(* IEC 61131-3 sources: JingjiangMoonbox/Application/Application/任务列表/TensionTask/张力控制/收放牵/张力控制, 5 files *)

(* ---- KS_FB_CalcGirthByVel_IfOf.st ---- *)
(*@CES
Name=KS_FB_CalcGirthByVel_IfOf
Type=FunctionBlock
TypeGuid=6f9dac99-8de1-4efc-8465-68ac443b7d08
Guid=2b108746-d302-40a1-8059-c5776d7629bb
HasDeclaration=True
HasImplementation=True
*)
{DECLARATION}
FUNCTION_BLOCK KS_FB_CalcGirthByVel_IfOf
VAR_INPUT
	i_xEn: BOOL;
	i_xCalcGirthEn:BOOL;(**)
	i_rVel_Film:REAL;(*料膜速度*)
	i_iCycleTime_Plc:INT;(*程序执行周期*)
	i_rAnalogLimit:REAL;(*模拟量的限值*)
	i_rUsingGirth:REAL;(*使用的周长值*)
	i_rAnalogSumLimit:REAL;(*模拟量累计值的限值*)
	i_rAxisVel_Cur:REAL;(*当前轴速度*)
	i_rAi_Swing: REAL; (*摆臂当前值*)
END_VAR
VAR_OUTPUT
	o_xEno:BOOL;
	o_iErNo: INT;
	o_xGirthCaled:BOOL;(*周长计算完成了~*)
	o_rGirth:REAL;(*计算出来的周长值*)
END_VAR
VAR
	rAver_CurrentVel: REAL;
	rCurrentVelSum:LREAL;(*当前速度累计值*)
	rAnalogSum: REAL; (*当前模拟量累计值*)
	iCycleCount: INT;
	arDataFifo:ARRAY [1..2,1..c_iArrNum] OF REAL;(*用来存放每个周期速度以及模拟量的值。一维数组代表速度值，二维数组代表模拟量值*)
	xArrInited: BOOL;		(*数组初始化完成*)
	iDelayCount: INT;
	iN: INT;
	xAnalogValue: BOOL;(*放牵模拟量有效*)
	iLastIndex: INT;
END_VAR
VAR CONSTANT
	c_iArrNum:INT:=300;(*数组大小暂定为100个 按20ms周期算就是2s的数据*)
								(*2019.7.25.125733 将计算周期拉长了！|Liu.yt*)
END_VAR
{IMPLEMENTATION}
o_xEno:= i_xEn;
o_iErNo:= 0;
IF i_xEn THEN

	o_xGirthCaled:=FALSE;(*该标志只有效一个周期*)
	o_rGirth:=0;
	rAver_CurrentVel:=0;
	rCurrentVelSum:=0;
	rAnalogSum:=0;

	IF i_xCalcGirthEn  THEN(*使能计算周长功能*)

		(*保存一定时间的速度值，用来进行平均速度计算。时间暂定为2s*)
		iCycleCount:=iCycleCount+1;(*计数+1*)
		IF iCycleCount>c_iArrNum THEN(*循环存储*)
			iCycleCount:=1;
		END_IF
		arDataFifo[1,iCycleCount]:=i_rAxisVel_Cur;(*速度值*)
		arDataFifo[2,iCycleCount]:=i_rAi_Swing;(*模拟量值*)

		(*周长计算*)
		IF iCycleCount>=c_iArrNum OR xArrInited THEN (*累计足够次数的速度值*)

			xArrInited:=TRUE;
			iDelayCount:=iDelayCount+1;
		(*计算模拟量累计值和速度累计值*)
			FOR iN:=1 TO c_iArrNum BY 1 DO
				rCurrentVelSum:=rCurrentVelSum+arDataFifo[1,iN];
				IF ABS(arDataFifo[2,iN])>i_rAnalogLimit AND iDelayCount<=500 THEN(*累计的这段时间里的模拟量值必须都小于等于模拟量限值才有效
												iDelayCount 是用来保证在极端情况下不能满足条件也可以进入计算逻辑*)
					rAnalogSum:=i_rAnalogSumLimit+1;(*给模拟量累计值一个大于模拟量累计限值的值，这样我们在下面的判断中则会认为无效*)
					xAnalogValue:=FALSE;
					EXIT;
				ELSE
					xAnalogValue:=TRUE;
					rAnalogSum:=rAnalogSum+arDataFifo[2,iN];
				END_IF
			END_FOR

			iLastIndex:=(iCycleCount+1) MOD c_iArrNum;

			IF ABS((arDataFifo[2,iCycleCount])-(arDataFifo[2,iLastIndex])) >0.005 OR NOT  xAnalogValue THEN(*模拟量2S的变化量超过范围，则认为无效*);
			ELSE(*模拟量累计值在一定范围内求取速度平均值*)
				rAver_CurrentVel:=rCurrentVelSum/INT_TO_REAL(c_iArrNum);
			END_IF
		END_IF

		IF rAver_CurrentVel<>0 AND i_rVel_Film<>0 THEN (*平均速度不等于0 我们认为已经计算出了满足条件的平均速度值*)
			o_rGirth:=i_rVel_Film*i_rUsingGirth/rAver_CurrentVel;(*计算出理论周长值*)
			o_xGirthCaled:=TRUE;
		END_IF
	ELSE
		iDelayCount:=0;
		iCycleCount:=0;
		xArrInited:=FALSE;
	END_IF
ELSE
	;
END_IF

(* ---- KS_FB_CalcGirthLogic_IfOf.st ---- *)
(*@CES
Name=KS_FB_CalcGirthLogic_IfOf
Type=FunctionBlock
TypeGuid=6f9dac99-8de1-4efc-8465-68ac443b7d08
Guid=2fd058fe-87b7-4e24-a0c2-a6df17a2c853
HasDeclaration=True
HasImplementation=True
*)
{DECLARATION}
FUNCTION_BLOCK KS_FB_CalcGirthLogic_IfOf
(*2021.10.28.100152 收放牵分开*)
(*默认调整方向|在摆臂越来越大时候即越来越紧|周长是加大方向也就是减速方向|
放牵调整方向需要取反|
收牵不需要*)
(*再切换算法后直接退出周长模式@2026.4.9.195445+*)
VAR_INPUT
	i_xEn:BOOL;
	i_xMachineRev:BOOL;(*反向走料时调整方向取反*)
	i_xNegative:BOOL;(*调整取反*)
	i_rVel_Film:REAL;(*当前料膜速度*)
	i_iCycleTime_Plc:INT;(*程序执行周期*)
	i_rAnalogLimit:REAL;(*模拟量有效值限值*)
	i_rAxisVel_Cur:REAL;(*当前轴速度*)
	i_rAi_Swing: REAL; (*摆臂当前值*)
	i_rActualGirth:REAL;(*默认周长*)
	i_xRollerPressDone: BOOL;
	i_xSwitchTension:BOOL;(*张力算法控制开关*)
	i_xAccing:BOOL;
	i_xDecing:BOOL;
	i_xCompensateWhenAccing:BOOL;(*2025.3.7.092457*)
	i_rCompensateGirthWhenAccing:REAL;(*补偿的值|mm*)
	i_iCycleNum_Delay: INT:= 500;
	i_iCycleNum_AI_Ave: INT:=50;
END_VAR
VAR_OUTPUT
	o_xEno: BOOL;
	o_iErNo: INT;
	o_xGirthCalFinish: BOOL;
	o_rUsingGirth: REAL;
END_VAR
VAR
	fbKS_FB_CalcGirthByVel: KS_FB_CalcGirthByVel_IfOf;
	xEvenning:BOOL;		(*稳速标志*)
	xAccing: BOOL;
	xDecing: BOOL;
	xConditionDone: BOOL;
	xCalGirthEn: BOOL;(*周长计算使能标志*)
	xGirthCaled:BOOL;(*计算好了*)
	xPreGirthCalFinish: BOOL;(*上个周期周长计算完成*)
	rGirthTemp: REAL;(*计算的周长值*)
	rPreCurVel: REAL;(*上个周期当前速度值*)
	iCalGirthCount: INT;(*周期计数值*)
	iGirthStep: INT:= 2;
	rGirthStep_Temp: REAL;
	iThreshold: INT:=5;(*计算出的的牵引周长有效范围单位%*)
	rAnalog_Sum: REAL;
	iCycleCount:INT;(*调整计时*)
	rAnalog_Aver:REAL;(*平均模拟量*)
	rPreAnalog_Aver: REAL;(*上次计算后的平均模拟量*)
	xCalAverDone: BOOL;(*平均值计算完成标志*)
	rThreshold: REAL;(*调整阈值*)
	iCoeff: INT;
	iCompensateGirthWhenAccing:INT;(*补偿的值|丝*)
END_VAR
VAR CONSTANT
	(*2020.4.22.101010_|新增|*)
	c_lrAIBoundage: LREAL := 0.5;
END_VAR
{IMPLEMENTATION}
o_xEno:= i_xEn;
o_iErNo:= 0;
IF i_xEn THEN
	(*稳速时候才能进行周长计算*)
	xEvenning:=NOT i_xAccing AND NOT i_xDecing AND i_rVel_Film>=9.9;(*编码器计算的速度,精度问题10m/min的时候回事9.99m/min*)
	xAccing:=i_xAccing;
	xDecing:=i_xDecing;

	xConditionDone:=FALSE;
	IF i_iCycleNum_Delay=0 THEN
		i_iCycleNum_Delay:= 500;
	END_IF
	IF xEvenning THEN(*进入匀速状态之后 等待一段时间在进入计算周长状态*)
		iCalGirthCount:=iCalGirthCount+1;
		IF iCalGirthCount>=i_iCycleNum_Delay THEN (*延迟500个周期 进入计算周长状态*)
			iCalGirthCount:=iCalGirthCount-1;
			xConditionDone:=TRUE;
		END_IF
	ELSE
		iCalGirthCount:=0;
	END_IF

	xCalGirthEn:=FALSE;
	IF xConditionDone AND NOT o_xGirthCalFinish  THEN
		xCalGirthEn:=TRUE;
	END_IF

	(*2018.08.16.81201 | niu.j |*)
	(*计算版周长使能取消，使用默认周长，一直调整*)
	IF i_xSwitchTension OR (NOT i_xRollerPressDone) THEN
		xCalGirthEn:= FALSE;
	END_IF
	(*------------------------------------------*)

	fbKS_FB_CalcGirthByVel(
		i_xEn:= TRUE,
		i_xCalcGirthEn:= xCalGirthEn,
		i_rVel_Film:= i_rVel_Film,
		i_iCycleTime_Plc:= i_iCycleTime_Plc,
		i_rAnalogLimit:= i_rAnalogLimit,
		i_rUsingGirth:= o_rUsingGirth,
		i_rAnalogSumLimit:= ,
		i_rAxisVel_Cur:= i_rAxisVel_Cur,
		i_rAi_Swing:= i_rAi_Swing,
		o_xEno=> ,
		o_xGirthCaled=> xGirthCaled,
		o_rGirth=> rGirthTemp);

	IF xGirthCaled THEN
		o_xGirthCalFinish:=TRUE;(*该标志有效则可以认为我们可以进入非调整状态了*)
	END_IF

	IF o_xGirthCalFinish AND ABS(i_rAi_Swing)>c_lrAIBoundage OR
		(NOT i_xRollerPressDone) OR(*2021.10.27.112505 压辊抬起来了就取消周长调整模式*)
		i_xSwitchTension THEN(*取消周长方式@直接进入pi方式@2026.3.18.140545+*)(*2026.4.9.194300同步*)
		o_xGirthCalFinish:=FALSE;
	END_IF

	IF o_xGirthCalFinish AND (NOT xPreGirthCalFinish) THEN(*将计算出来的值赋给输出值*)
		IF rGirthTemp<=i_rActualGirth*(1+iThreshold/100.0) AND rGirthTemp>=i_rActualGirth*(1-iThreshold/100.0) THEN
			o_rUsingGirth:=rGirthTemp;
		ELSE
			o_xGirthCalFinish:=FALSE;
		END_IF
	END_IF

	IF i_rVel_Film<=0.01 THEN(*不走料的时候版周长为默认值*)
		o_xGirthCalFinish:=FALSE;
		o_rUsingGirth:= i_rActualGirth;
	END_IF

	(*当已经进入到不再调整逻辑中的时候，我们对牵引的周长进行微调*)(*2018.5.7.153458*)

	(*求摆臂的位置的平均值*)
	xCalAverDone:=FALSE;
	iCycleCount:=iCycleCount+1;
	rAnalog_Sum:=rAnalog_Sum+i_rAi_Swing;
	IF i_iCycleNum_AI_Ave=0 THEN
		i_iCycleNum_AI_Ave:= 50;
	END_IF
	IF iCycleCount>=i_iCycleNum_AI_Ave THEN
		xCalAverDone:=TRUE;
		rAnalog_Aver:=rAnalog_Sum/iCycleCount;
		rAnalog_Sum:=0;
		iCycleCount:=0;
	ELSE;
	END_IF

	IF o_xGirthCalFinish AND NOT xPreGirthCalFinish  THEN(*计算完成后初始化上个周期平均模拟量值*)
		rPreAnalog_Aver:=rAnalog_Aver;
	END_IF

	rGirthTemp:=0;
(*2022.8.11.093253更新版周长调整当量--变速时是2丝--稳速1丝||liu&chen&niu*)
	IF xEvenning THEN
		rGirthStep_Temp:= 1;
	ELSIF (xDecing OR xAccing) AND i_rVel_Film>=10 THEN
		rGirthStep_Temp:= INT_TO_REAL(iGirthStep);
	ELSE
		rGirthStep_Temp:= 1;
	END_IF

	rGirthStep_Temp:=rGirthStep_Temp/100.0;
	IF o_xGirthCalFinish AND xCalAverDone  THEN
		IF ABS(rAnalog_Aver)>0.1 THEN
			rThreshold:=0;
		ELSE
			rThreshold:=0.001;
		END_IF

		IF NOT i_xMachineRev THEN
			iCoeff:=1;
		ELSE
			iCoeff:=-1;
		END_IF
		(*调整取反|同样变化趋势补偿方向不同*)
		IF i_xNegative THEN
			iCoeff:=-iCoeff;
		END_IF

		IF  rAnalog_Aver >0.01 THEN
			IF  rAnalog_Aver>rPreAnalog_Aver+rThreshold THEN(*位置值越来越大了*)
				rGirthTemp:=iCoeff*rGirthStep_Temp;
				rPreAnalog_Aver:=rAnalog_Aver;
			END_IF
		ELSIF  rAnalog_Aver <-0.01  THEN
			IF  rAnalog_Aver+rThreshold<rPreAnalog_Aver THEN(*位置值越来越小了*)
				rGirthTemp:=-iCoeff*rGirthStep_Temp;
				rPreAnalog_Aver:=rAnalog_Aver;
			END_IF
		ELSE
			rPreAnalog_Aver:=rAnalog_Aver;
		END_IF
	ELSE;
	END_IF
	(*放料升速开始周长补偿值处理*)
	IF i_xAccing THEN
		IF i_xCompensateWhenAccing THEN
			IF iCompensateGirthWhenAccing>0 THEN
				IF iCompensateGirthWhenAccing-rGirthStep_Temp*100<0 THEN
					rGirthTemp:=rGirthTemp+INT_TO_REAL(iCompensateGirthWhenAccing)/100;
					iCompensateGirthWhenAccing:=0;
				ELSE
					rGirthTemp:=rGirthTemp+rGirthStep_Temp;
					iCompensateGirthWhenAccing:=LREAL_TO_INT(iCompensateGirthWhenAccing-rGirthStep_Temp*100);
				END_IF
			ELSIF iCompensateGirthWhenAccing<0 THEN
				IF iCompensateGirthWhenAccing+rGirthStep_Temp*100>0 THEN
					rGirthTemp:=rGirthTemp-INT_TO_REAL(iCompensateGirthWhenAccing)/100;
					iCompensateGirthWhenAccing:=0;
				ELSE
					rGirthTemp:=rGirthTemp-rGirthStep_Temp;
					iCompensateGirthWhenAccing:=LREAL_TO_INT(iCompensateGirthWhenAccing+rGirthStep_Temp*100);
				END_IF
			ELSE;
			END_IF
		END_IF
	ELSE
		iCompensateGirthWhenAccing:=REAL_TO_INT(i_rCompensateGirthWhenAccing*100);
	END_IF

	o_rUsingGirth:=o_rUsingGirth+rGirthTemp;

	rPreCurVel:=i_rVel_Film;
	xPreGirthCalFinish:=o_xGirthCalFinish;
ELSE
	IF o_rUsingGirth=0 THEN
		o_rUsingGirth:= i_rActualGirth;
	END_IF
END_IF

(* ---- KS_FB_CalcGirthLogic_IfOf_BAK.st ---- *)
(*@CES
Name=KS_FB_CalcGirthLogic_IfOf_BAK
Type=FunctionBlock
TypeGuid=6f9dac99-8de1-4efc-8465-68ac443b7d08
Guid=07fd00ea-7360-439f-a038-63e58a6ffd7e
HasDeclaration=True
HasImplementation=True
*)
{DECLARATION}
FUNCTION_BLOCK KS_FB_CalcGirthLogic_IfOf_BAK
(*2021.10.28.100152 收放牵分开*)
(*默认调整方向|在摆臂越来越大时候即越来越紧|周长是加大方向也就是减速方向|
放牵调整方向需要取反|
收牵不需要*)
VAR_INPUT
	i_xEn:BOOL;
	i_xMachineRev:BOOL;(*反向走料时调整方向取反*)
	i_xNegative:BOOL;(*调整取反*)
	i_rVel_Film:REAL;(*当前料膜速度*)
	i_iCycleTime_Plc:INT;(*程序执行周期*)
	i_rAnalogLimit:REAL;(*模拟量有效值限值*)
	i_rAxisVel_Cur:REAL;(*当前轴速度*)
	i_rAi_Swing: REAL; (*摆臂当前值*)
	i_rActualGirth:REAL;(*默认周长*)
	i_xRollerPressDone: BOOL;
	i_xSwitchTension:BOOL;(*张力算法控制开关*)
	i_xAccing:BOOL;
	i_xDecing:BOOL;
	i_xCompensateWhenAccing:BOOL;(*2025.3.7.092457*)
	i_rCompensateGirthWhenAccing:REAL;(*补偿的值|mm*)
	i_iCycleNum_Delay: INT:= 500;
	i_iCycleNum_AI_Ave: INT:=50;
END_VAR
VAR_OUTPUT
	o_xEno: BOOL;
	o_iErNo: INT;
	o_xGirthCalFinish: BOOL;
	o_rUsingGirth: REAL;
END_VAR
VAR
	fbKS_FB_CalcGirthByVel: KS_FB_CalcGirthByVel_IfOf;
	xEvenning:BOOL;		(*稳速标志*)
	xAccing: BOOL;
	xDecing: BOOL;
	xConditionDone: BOOL;
	xCalGirthEn: BOOL;(*周长计算使能标志*)
	xGirthCaled:BOOL;(*计算好了*)
	xPreGirthCalFinish: BOOL;(*上个周期周长计算完成*)
	rGirthTemp: REAL;(*计算的周长值*)
	rPreCurVel: REAL;(*上个周期当前速度值*)
	iCalGirthCount: INT;(*周期计数值*)
	iGirthStep: INT:= 2;
	rGirthStep_Temp: REAL;
	iThreshold: INT:=5;(*计算出的的牵引周长有效范围单位%*)
	rAnalog_Sum: REAL;
	iCycleCount:INT;(*调整计时*)
	rAnalog_Aver:REAL;(*平均模拟量*)
	rPreAnalog_Aver: REAL;(*上次计算后的平均模拟量*)
	xCalAverDone: BOOL;(*平均值计算完成标志*)
	rThreshold: REAL;(*调整阈值*)
	iCoeff: INT;
	iCompensateGirthWhenAccing:INT;(*补偿的值|丝*)
END_VAR
VAR CONSTANT
	(*2020.4.22.101010_|新增|*)
	c_lrAIBoundage: LREAL := 0.5;
END_VAR
{IMPLEMENTATION}
o_xEno:= i_xEn;
o_iErNo:= 0;
IF i_xEn THEN
	(*稳速时候才能进行周长计算*)
	xEvenning:=NOT i_xAccing AND NOT i_xDecing AND i_rVel_Film>=10;
	xAccing:=i_xAccing;
	xDecing:=i_xDecing;

	xConditionDone:=FALSE;
	IF i_iCycleNum_Delay=0 THEN
		i_iCycleNum_Delay:= 500;
	END_IF
	IF xEvenning THEN(*进入匀速状态之后 等待一段时间在进入计算周长状态*)
		iCalGirthCount:=iCalGirthCount+1;
		IF iCalGirthCount>=i_iCycleNum_Delay THEN (*延迟500个周期 进入计算周长状态*)
			iCalGirthCount:=iCalGirthCount-1;
			xConditionDone:=TRUE;
		END_IF
	ELSE
		iCalGirthCount:=0;
	END_IF

	xCalGirthEn:=FALSE;
	IF xConditionDone AND NOT o_xGirthCalFinish  THEN
		xCalGirthEn:=TRUE;
	END_IF

	(*2018.08.16.81201 | niu.j |*)
	(*计算版周长使能取消，使用默认周长，一直调整*)
	IF i_xSwitchTension OR (NOT i_xRollerPressDone) THEN
		xCalGirthEn:= FALSE;
	END_IF
	(*------------------------------------------*)

	fbKS_FB_CalcGirthByVel(
		i_xEn:= TRUE,
		i_xCalcGirthEn:= xCalGirthEn,
		i_rVel_Film:= i_rVel_Film,
		i_iCycleTime_Plc:= i_iCycleTime_Plc,
		i_rAnalogLimit:= i_rAnalogLimit,
		i_rUsingGirth:= o_rUsingGirth,
		i_rAnalogSumLimit:= ,
		i_rAxisVel_Cur:= i_rAxisVel_Cur,
		i_rAi_Swing:= i_rAi_Swing,
		o_xEno=> ,
		o_xGirthCaled=> xGirthCaled,
		o_rGirth=> rGirthTemp);

	IF xGirthCaled THEN
		o_xGirthCalFinish:=TRUE;(*该标志有效则可以认为我们可以进入非调整状态了*)
	END_IF

	IF o_xGirthCalFinish AND ABS(i_rAi_Swing)>c_lrAIBoundage OR
		(NOT i_xRollerPressDone) THEN(*2021.10.27.112505 压辊抬起来了就取消周长调整模式*)
		o_xGirthCalFinish:=FALSE;
	END_IF

	IF o_xGirthCalFinish AND (NOT xPreGirthCalFinish) THEN(*将计算出来的值赋给输出值*)
		IF rGirthTemp<=i_rActualGirth*(1+iThreshold/100.0) AND rGirthTemp>=i_rActualGirth*(1-iThreshold/100.0) THEN
			o_rUsingGirth:=rGirthTemp;
		ELSE
			o_xGirthCalFinish:=FALSE;
		END_IF
	END_IF

	IF i_rVel_Film<=0.01 THEN(*不走料的时候版周长为默认值*)
		o_xGirthCalFinish:=FALSE;
		o_rUsingGirth:= i_rActualGirth;
	END_IF

	(*当已经进入到不再调整逻辑中的时候，我们对牵引的周长进行微调*)(*2018.5.7.153458*)

	(*求摆臂的位置的平均值*)
	xCalAverDone:=FALSE;
	iCycleCount:=iCycleCount+1;
	rAnalog_Sum:=rAnalog_Sum+i_rAi_Swing;
	IF i_iCycleNum_AI_Ave=0 THEN
		i_iCycleNum_AI_Ave:= 50;
	END_IF
	IF iCycleCount>=i_iCycleNum_AI_Ave THEN
		xCalAverDone:=TRUE;
		rAnalog_Aver:=rAnalog_Sum/iCycleCount;
		rAnalog_Sum:=0;
		iCycleCount:=0;
	ELSE;
	END_IF

	IF o_xGirthCalFinish AND NOT xPreGirthCalFinish  THEN(*计算完成后初始化上个周期平均模拟量值*)
		rPreAnalog_Aver:=rAnalog_Aver;
	END_IF

	rGirthTemp:=0;
(*2022.8.11.093253更新版周长调整当量--变速时是2丝--稳速1丝||liu&chen&niu*)
	IF xEvenning THEN
		rGirthStep_Temp:= 1;
	ELSIF (xDecing OR xAccing) AND i_rVel_Film>=10 THEN
		rGirthStep_Temp:= INT_TO_REAL(iGirthStep);
	ELSE
		rGirthStep_Temp:= 1;
	END_IF

	rGirthStep_Temp:=rGirthStep_Temp/100.0;
	IF o_xGirthCalFinish AND xCalAverDone  THEN
		IF ABS(rAnalog_Aver)>0.1 THEN
			rThreshold:=0;
		ELSE
			rThreshold:=0.001;
		END_IF

		IF NOT i_xMachineRev THEN
			iCoeff:=1;
		ELSE
			iCoeff:=-1;
		END_IF
		(*调整取反|同样变化趋势补偿方向不同*)
		IF i_xNegative THEN
			iCoeff:=-iCoeff;
		END_IF

		IF  rAnalog_Aver >0.01 THEN
			IF  rAnalog_Aver>rPreAnalog_Aver+rThreshold THEN(*位置值越来越大了*)
				rGirthTemp:=iCoeff*rGirthStep_Temp;
				rPreAnalog_Aver:=rAnalog_Aver;
			END_IF
		ELSIF  rAnalog_Aver <-0.01  THEN
			IF  rAnalog_Aver+rThreshold<rPreAnalog_Aver THEN(*位置值越来越小了*)
				rGirthTemp:=-iCoeff*rGirthStep_Temp;
				rPreAnalog_Aver:=rAnalog_Aver;
			END_IF
		ELSE
			rPreAnalog_Aver:=rAnalog_Aver;
		END_IF
	ELSE;
	END_IF
	(*放料升速开始周长补偿值处理*)
	IF i_xAccing THEN
		IF i_xCompensateWhenAccing THEN
			IF iCompensateGirthWhenAccing>0 THEN
				IF iCompensateGirthWhenAccing-rGirthStep_Temp*100<0 THEN
					rGirthTemp:=rGirthTemp+INT_TO_REAL(iCompensateGirthWhenAccing)/100;
					iCompensateGirthWhenAccing:=0;
				ELSE
					rGirthTemp:=rGirthTemp+rGirthStep_Temp;
					iCompensateGirthWhenAccing:=LREAL_TO_INT(iCompensateGirthWhenAccing-rGirthStep_Temp*100);
				END_IF
			ELSIF iCompensateGirthWhenAccing<0 THEN
				IF iCompensateGirthWhenAccing+rGirthStep_Temp*100>0 THEN
					rGirthTemp:=rGirthTemp-INT_TO_REAL(iCompensateGirthWhenAccing)/100;
					iCompensateGirthWhenAccing:=0;
				ELSE
					rGirthTemp:=rGirthTemp-rGirthStep_Temp;
					iCompensateGirthWhenAccing:=LREAL_TO_INT(iCompensateGirthWhenAccing+rGirthStep_Temp*100);
				END_IF
			ELSE;
			END_IF
		END_IF
	ELSE
		iCompensateGirthWhenAccing:=REAL_TO_INT(i_rCompensateGirthWhenAccing*100);
	END_IF

	o_rUsingGirth:=o_rUsingGirth+rGirthTemp;

	rPreCurVel:=i_rVel_Film;
	xPreGirthCalFinish:=o_xGirthCalFinish;
ELSE
	IF o_rUsingGirth=0 THEN
		o_rUsingGirth:= i_rActualGirth;
	END_IF
END_IF

(* ---- KS_FB_TensionCtl_IfOf.st ---- *)
(*@CES
Name=KS_FB_TensionCtl_IfOf
Type=FunctionBlock
TypeGuid=6f9dac99-8de1-4efc-8465-68ac443b7d08
Guid=b7b8bc31-4f35-42b3-88de-f6b214f8ce5f
HasDeclaration=True
HasImplementation=True
*)
{DECLARATION}
FUNCTION_BLOCK KS_FB_TensionCtl_IfOf
(*摆臂负值-料膜为松弛状态|负值输出减速|反之加速*)
(*2021.10.23.093343  新增的张力控制模块|主要用于收放牵控制*)
VAR_INPUT
	i_xEn: BOOL;(*张力模块使能*)
	i_xCanAdjEn: BOOL;(*调整和非调整切换标志|算法需要*)
	i_xIsDebugMode:BOOL;(*调试模式*)
	i_xNegative_PiValue:BOOL;(*pi取反*)
	i_xMachineRev:BOOL;(*反向走料信号*)
	i_rAI_Swing: REAL; (*摆臂模拟量*)
	i_rVel_Film:REAL;(*当前料膜速度*)
//	i_iPiVelLimit:INT;(*pi限值-最大调整10M/MIN*)
	i_xFilmAccDecDone:BOOL;(*料膜加速完成标志*)
	i_iTimeTo0WhenDisEn:INT:=1;(*当前速度在取消使能时到0速的规划时间|s-写0则不规划*)
	i_iCycleTime_Plc:INT;(*程序执行周期*)
	i_rKp:REAL;
	i_rKi:REAL;
	i_rKd:REAL;
	i_byVelLimit_PerCent:BYTE;(*速度限制百分比%*)
	i_xFeedlimitWarnFlag:BOOL;(*牵引速度限制提示开关*)
	i_iFeedLimitWarnCoff: INT;(*牵引限制系数*)
	i_rUsingGirth:REAL;(*调整后的周长返回值*)
	i_xAdjustMode:BOOL;(*调整开关*)
	i_rGirth_Input:REAL;(*界面输入周长*)
	i_iVel_Max:INT;(*主机最大速度|2021.2.2.110402 增加|调整else的时候使用最大速度计算加速度*)

	i_uiMaxVel_UseCalcAcc:UINT;(*最大速度,用于计算最大加减速@2024.04.12.165352*)

	(*2024.05.24.110325+*)
	i_xPseudoRandomId					:BOOL;(*=True*)
	i_xPseudoRandomEn					:BOOL;(*伪随机使能|功能使能*)
	i_xPseudoRandomTsting				:BOOL;(*伪随机使能了*)
	i_rPseudoRandomRoundAmplitude_Cur	:REAL;
	i_pbySetTestPid						:POINTER TO BYTE;(*设置测试的pid*)
	i_iPseudoRandomRound_Kp_1			:INT;
	i_iPseudoRandomRound_Kd_1			:INT;
	i_iPseudoRandomRound_Kp_2			:INT;
	i_iPseudoRandomRound_Kd_2			:INT;
	i_iPseudoRandomRound_Kp_3			:INT;
	i_iPseudoRandomRound_Kd_3			:INT;

	i_xPidType						:BOOL;(*false=原来方式\true=新的*)

	i_xUseAntiNotch					:BOOL;(*输入使用陷波*)
	i_prWn							:POINTER TO REAL;
	i_prBw							:POINTER TO REAL;
	i_prDp							:POINTER TO REAL;

	(*扰动输出的控制输入参数@2024.12.3.102359*)
	i_xEn_Disturbance:BOOL;(*扰动使能@需要常有效*)
	i_rFreq_Disturbance:REAL;(*扰动频率@hz*)
	i_rAmplitude_Disturbance:REAL;(*扰动幅值*)
	i_uiTotalTime_Disturbance:UINT;(*扰动输出的总时间|=0 代表一直输出@s*)

	i_xRollerSts_Pu: BOOL;
END_VAR
VAR_OUTPUT
	o_xEno :BOOL;
	o_iErNo: INT;
	o_rVel: REAL;
	o_rPi_Value:REAL;
	o_rForwardStep:REAL;
	o_rVel_rpm:REAL;(*转速@r/min*)
	o_xOuting_sin:BOOL;(*正弦输出中@2024.12.3.110839*)
	o_rResult_sin:REAL;(*正弦输出值@2024.12.3.110839*)
END_VAR
VAR
	iN: INT;
	rKp : REAL; (*P值*)
	rKi : REAL; (*I值*)
	rKd: REAL;(*D值*)

	iVoltTotalTimes: INT := 0;
	iVoltAverageMaxTimes: INT := 20; (*模拟采集平均次数*)
	arVolt: ARRAY [1..20] OF REAL := [20(0)]; (*历史模拟量列表*)
	rVoltSum: REAL; (*模拟量累计*)
	rFormulaResult: REAL; (*PID运算后的放牵调整值*)
	rVoltFinal: REAL; (*最终用的模拟量*)
	rTempResult: REAL; (*临时的输出结果*)
	rMaxDelVel: REAL;
	rForwardStep: REAL;(*前馈步进值*)
	rPreFilmVelocity: REAL;
	rPIValueLimit_Zero: REAL:=0.02;(*0速最大调整量*)
	iVelocityLimit: INT:=2;(*零速最大调整速度限值*)
	iNum_Old: INT := 5;
	iTimeTo0WhenDisEn:INT:=1;(*当前速度在取消使能时到0速的规划时间|s*)
	lrVel_Acceleration: LREAL:=0;(*速度规划到0加速度*)
	xFilmDecFlag: BOOL:=FALSE;(*料膜减速标志*)
	rTempVel: REAL;(*临时速度*)
	xIsDebugging: BOOL;(*调试中标志*)
	arAntiNotchU_Uk: ARRAY [1..3] OF REAL;
	arAntiNotchU_Yk: ARRAY [1..3] OF REAL;
	rAntiNotch_Out: REAL;
	rAI_cur: REAL;
	bySetTestPid: BYTE;(*设置伪随机pid*)
	rDeltaTmp: REAL;
	rPseudoRandomRoundAmplitude_Cur: REAL;(*伪随机当前值*)
	rPseudoRandomRoundAmplitude_Cur_Last: REAL;
	rPseudoRandomAmplitude_Delta: REAL;
	(*2024.05.25.104740*)
	rYI: REAL;(*积分控制输出寄存器*)
	rYD: REAL;(*微分控制输出寄存器*)
	rYout: REAL;
	arEk:ARRAY [1..2] OF REAL;(*误差寄存器 [e(k);e(k-1)]*)
	(*2025.1.12.152712+*)
	rYout_Tmp: REAL;
	xCtlEn: BOOL;(*控制使能*)
	xCtlEn_Last: BOOL;
	lrX_sin:LREAL;(*正弦的时间轴*)
	rResult_sin:REAL;(*正弦值*)
	rVel_Disturbance: REAL;(*放牵扰动值*)
	rTmp: REAL;
	rDelt: REAL;
	lrTempVel: LREAL;
END_VAR
{IMPLEMENTATION}
rMaxDelVel:=0.3;(*=300/20/50 20S加速到300m/min的时候一个周期速度的变化量*)(*2018.5.22.115216 增加调整量限值*)
rPIValueLimit_Zero:=0.03;(*0速时调整量限值*)
//iVelocityLimit:=i_iPiVelLimit;

(*2022.9.20.143232 速度限制使用%|最小2m/min 最大10m/min*)
IF i_byVelLimit_PerCent<>0 THEN
	iVelocityLimit:=LREAL_TO_INT(i_byVelLimit_PerCent*i_rVel_Film/100);
ELSE(*等于0按照10m/min限制-以前一直使用该值*)
	iVelocityLimit:=10;
END_IF

IF iVelocityLimit<2 THEN
	iVelocityLimit:=2;
ELSIF iVelocityLimit>10 THEN
	iVelocityLimit:=10;
END_IF

IF i_rVel_Film=0 THEN(*料膜速度为0速的时候，调整牵引到中位。对速度进行限值*)(*2018.7.11.223054*)
	iVelocityLimit:=2;
END_IF
(*2025.3.7.100539*)
(*参数初始化*)
IF i_prWn<>0 AND i_prBw<>0 AND i_prDp <>0 THEN
	IF i_prWn^=0 THEN
		i_prWn^:=1;
	END_IF
	IF i_prBw^=0 THEN
		i_prBw^:=2;
	END_IF
	IF i_prDp^=0 THEN
		i_prDp^:=20;
	END_IF
END_IF

IF i_xEn AND i_rVel_Film>0 THEN
	(*放牵*)
	IF i_prWn<>0 AND i_prBw<>0 AND i_prDp <>0 THEN
		AntiNotch(
			i_rAI_Swing(*i_rU*),
			ADR(rAntiNotch_Out)(*i_prYout*),
			i_prWn^(*i_rWn*),
			i_prBw^(*i_rBw*),
			i_prDp^(*i_rDp*),
			INT_TO_REAL(i_iCycleTime_Plc)/1000.0(*i_rTs*),
			ADR(arAntiNotchU_Uk)(*i_prUk*),
			ADR(arAntiNotchU_Yk)(*i_prYk*));
	END_IF
ELSE
	SysMemSet(ADR(arAntiNotchU_Uk),0,SIZEOF(arAntiNotchU_Uk));
	SysMemSet(ADR(arAntiNotchU_Yk),0,SIZEOF(arAntiNotchU_Yk));
END_IF

IF i_xUseAntiNotch THEN
	rAI_cur:=rAntiNotch_Out;
ELSE
	rAI_cur:=i_rAI_Swing;
END_IF

(*han.dp@2017-08-13 15:49:11
/.重新对要使用的模拟量进行一个简单的滤波
/.*)
FOR iN:=iVoltAverageMaxTimes TO 2 BY -1 DO
	arVolt[iN]:= arVolt[iN-1];
END_FOR
arVolt[1]:= rAI_cur;

(*求累计*)
rVoltSum:= 0;
FOR iN:=iVoltAverageMaxTimes TO 1 BY -1 DO
	rVoltSum:= rVoltSum + arVolt[iN];
END_FOR

IF iVoltTotalTimes<iVoltAverageMaxTimes THEN
	(*不足平均的次数就去当前值*)
	iVoltTotalTimes:= iVoltTotalTimes+1;
	rVoltFinal:= arVolt[1];
ELSE
	(*取平均值*)
	rVoltFinal:= rVoltSum/iVoltAverageMaxTimes;
END_IF

(*伪随机测试@2024.05.24.130600*)
(*PID值处理---------------------------------------start*)
IF i_pbySetTestPid<>0 THEN
	bySetTestPid:=i_pbySetTestPid^;
END_IF
IF i_xPseudoRandomId THEN(*收牵伪随机*)
	IF i_xPseudoRandomEn THEN(*伪随机使能了*)
		(*pid界面按钮修改*)
		IF bySetTestPid=1 THEN(*第一组pid*)
			IF i_xPseudoRandomId THEN(*放牵伪随机*)
				rKp:=i_iPseudoRandomRound_Kp_1;
				rKd:=i_iPseudoRandomRound_Kd_1;
			END_IF
		ELSIF bySetTestPid=2 THEN(*第二组pid*)
			IF i_xPseudoRandomId THEN(*放牵伪随机*)
				rKp:=i_iPseudoRandomRound_Kp_2;
				rKd:=i_iPseudoRandomRound_Kd_2;
			END_IF
		ELSIF bySetTestPid=3 THEN(*第三组pid*)
			IF i_xPseudoRandomId THEN(*放牵伪随机*)
				rKp:=i_iPseudoRandomRound_Kp_3;
				rKd:=i_iPseudoRandomRound_Kd_3;
			END_IF
		ELSIF bySetTestPid=4 THEN(*第4组pid@0*)
			IF i_xPseudoRandomId THEN(*放牵伪随机*)
				rKp:=0;
				rKd:=0;
			END_IF
		END_IF
	END_IF
END_IF
bySetTestPid:=0;

(*非伪随机\使用界面pid@2024.05.24.112400*)
IF (NOT i_xPseudoRandomId) OR(*未选择牵引*)
	(NOT i_xPseudoRandomEn) THEN(*未使能*)
	rKp:= i_rKp;
	rKi:= i_rKi;
	rKd:= i_rKd;
END_IF

IF i_pbySetTestPid<>0 THEN
	i_pbySetTestPid^:=bySetTestPid;
END_IF
(*PID值处理---------------------------------------end*)

(*伪随机值处理------------------------------------start*)
(*取变化的增量值*)
IF i_xPseudoRandomId THEN(*伪随机*)
	rPseudoRandomRoundAmplitude_Cur:=i_rPseudoRandomRoundAmplitude_Cur;
ELSE
	rPseudoRandomRoundAmplitude_Cur:=0;
END_IF
rDeltaTmp:=rPseudoRandomRoundAmplitude_Cur-rPseudoRandomRoundAmplitude_Cur_Last;
rPseudoRandomRoundAmplitude_Cur_Last:=rPseudoRandomRoundAmplitude_Cur;

rPseudoRandomAmplitude_Delta:=0;
IF i_xPseudoRandomTsting THEN(*伪随机中*)
	IF i_xPseudoRandomId THEN(*放牵*)
		rPseudoRandomAmplitude_Delta:=rDeltaTmp;
	END_IF
ELSE
	IF rDeltaTmp<>0 THEN
		IF i_xPseudoRandomId THEN(*放牵*)
			rPseudoRandomAmplitude_Delta:=rDeltaTmp;
		END_IF
	END_IF
END_IF

(*2024.05.25.105317*)
xCtlEn:=i_xEn AND i_rVel_Film>0;
IF (xCtlEn AND NOT xCtlEn_Last)THEN(*初始化*)
	rYout:=0;
	rYout_Tmp:=0;
	rYI:=0;
	rYD:=0;
	SysMemSet(ADR(arEk),0,SIZEOF(arEk));
END_IF
xCtlEn_Last:=xCtlEn;

(*放牵pid*)
PID_ANTI(
	rAI_cur(*i_rU*),
	(*调整量使用临时值处理@2025.1.12.152843*)
	ADR(rYout_Tmp)(*i_prYout*),
	rKp*6.3/30(*i_rP*),
	rKI*7/50(*i_rI*),
	0(*i_rD*),
	0(*i_rN*),
	INT_TO_REAL(i_iCycleTime_Plc)/1000.0(*i_rTs*),
	INT_TO_REAL(iVelocityLimit)(*i_rLim*),
	1(*i_rAntiWindup*),
	ADR(rYI)(*i_prYI*),
	ADR(rYD)(*i_prYD*),
	ADR(arEk)(*i_parEk*));
(*对调整量输出做平滑处理@变化增加限值*)
rYout:=KS_A2B_SmoothDeal(rYout,rYout_Tmp,rMaxDelVel);

(*2024.12.3.110816+*)
KS_SIG_SIN(
	i_xEn_Disturbance(*i_xEn*),
	i_rFreq_Disturbance(*i_rFreq*),
	i_rAmplitude_Disturbance(*i_rAmplitude*),
	i_uiTotalTime_Disturbance(*i_uiTotalTime*),
	i_iCycleTime_Plc(*i_iCycleTime_Plc*),
	ADR(o_xOuting_sin)(*i_pxOuting*),
	ADR(lrX_sin)(*i_plrX*),
	ADR(o_rResult_sin)(*i_prResult*));

rVel_Disturbance:=o_rResult_sin;
IF NOT i_xAdjustMode OR(*放牵周长调整方式下|不能叠加扰动*)
	NOT i_xCanAdjEn OR(*放牵未pid调整*)
	NOT xCtlEn THEN(*未使能也先清除了吧*)
	rVel_Disturbance:=0;
END_IF

IF xCtlEn(*i_xEn AND i_lrVel_Film>0*) THEN(*2024.05.25.105235*)
	rForwardStep:=0;
	IF i_xFilmAccDecDone THEN(*料膜加速完成了，才使用前馈*)
		IF i_rVel_Film<>rPreFilmVelocity AND rPreFilmVelocity<>0  THEN (*速度发生了变化*)
			rForwardStep:=(i_rVel_Film-rPreFilmVelocity);
		ELSE;
		END_IF
	END_IF

	IF NOT i_xMachineRev THEN
	(*放牵速度控制*)
		IF i_xCanAdjEn (*AND i_xImpressFlag_Pu*) THEN (*放牵合压*)
							(*2018.10.6.122439 取消色组压辊合压放牵才调整逻辑by liu.yt*)

			rFormulaResult:= rKp * rAI_cur/1000 +rKd/100*(arVolt[1]-arVolt[iNum_Old]); (*/100是为了输入Kp和Ki时放大了100倍*)
			IF  ABS(rFormulaResult)>rMaxDelVel THEN
				rFormulaResult:=rMaxDelVel*(rFormulaResult)/ABS(rFormulaResult);
			ELSE
				;
			END_IF

			IF i_rVel_Film=0 THEN(*料膜速度为0速的时候，调整牵引到中位。对pi调整量进行限值*)(*2018.7.11.223054*)
				IF ABS(rFormulaResult)>rPIValueLimit_Zero THEN
					rFormulaResult:=rPIValueLimit_Zero*rFormulaResult/ABS(rFormulaResult);
				END_IF
			END_IF

			(*pi输出取反*)
			IF i_xNegative_PiValue THEN
				rFormulaResult:=-rFormulaResult;
			END_IF

			IF o_rVel+rFormulaResult+rForwardStep<0 THEN
				IF i_rVel_Film=0 THEN
					o_rVel:=o_rVel+rFormulaResult+rForwardStep;
				ELSE
					o_rVel:=0;
				END_IF
			ELSE
				o_rVel:=o_rVel+rFormulaResult+rForwardStep;
			END_IF

			IF i_xCanAdjEn THEN (*调整标志有效*);
			ELSE(*不调整状态*)
				o_rVel:=i_rVel_Film;
			END_IF

	(*对输出的收放牵速度进行限值*)
			IF o_rVel >INT_TO_REAL(iVelocityLimit)+i_rVel_Film THEN
				o_rVel:=INT_TO_REAL(iVelocityLimit)+i_rVel_Film ;
			ELSIF o_rVel <-INT_TO_REAL(iVelocityLimit)+i_rVel_Film  THEN
				o_rVel:=-INT_TO_REAL(iVelocityLimit)+i_rVel_Film ;
			ELSE
				;
			END_IF
		ELSE
			o_rVel:=i_rVel_Film;
		END_IF
	ELSE(*反向走料调整取反*)
		IF i_xCanAdjEn AND i_xRollerSts_Pu THEN (*放牵合压*)
							(*2018.10.6.122439 取消色组压辊合压放牵才调整逻辑by liu.yt*)

			rFormulaResult:= rKp * (-rAI_cur)/1000 -rKd/100*(arVolt[1]-arVolt[iNum_Old]); (*/100是为了输入Kp和Ki时放大了100倍*)
	(*	lrFeedPI_Value:=i_lrFeed_lrP/1000*(i_Analog.lrAnalogInput_Feed)+i_lrFeed_lrD/100*(lrFeed_Voltage_Sum[1]-lrFeed_Voltage_Sum[iNum_Old]);*)

			IF  ABS(rFormulaResult)>rMaxDelVel THEN
				rFormulaResult:=rMaxDelVel*(rFormulaResult)/ABS(rFormulaResult);
			ELSE
				;
			END_IF

			IF i_rVel_Film=0 THEN(*料膜速度为0速的时候，调整牵引到中位。对pi调整量进行限值*)(*2018.7.11.223054*)
				IF ABS(rFormulaResult)>rPIValueLimit_Zero THEN
					rFormulaResult:=rPIValueLimit_Zero*rFormulaResult/ABS(rFormulaResult);
				END_IF
			END_IF

			(*pi输出取反*)
			IF i_xNegative_PiValue THEN
				rFormulaResult:=-rFormulaResult;
			END_IF

			IF o_rVel+rFormulaResult+rForwardStep<0 THEN
				IF i_rVel_Film=0 THEN
					o_rVel:=o_rVel+rFormulaResult+rForwardStep;
				ELSE
					o_rVel:=0;
				END_IF
			ELSE
				o_rVel:=o_rVel+rFormulaResult+rForwardStep;
			END_IF

			IF i_xCanAdjEn THEN (*调整标志有效*)
				;
			ELSE(*不调整状态*)
				o_rVel:=i_rVel_Film;
			END_IF

	(*对输出的收放牵速度进行限值*)
			IF o_rVel >INT_TO_REAL(iVelocityLimit)+i_rVel_Film THEN
				o_rVel:=INT_TO_REAL(iVelocityLimit)+i_rVel_Film ;
			ELSIF o_rVel <-INT_TO_REAL(iVelocityLimit)+i_rVel_Film  THEN
				o_rVel:=-INT_TO_REAL(iVelocityLimit)+i_rVel_Film ;
			ELSE
				;
			END_IF
		ELSE
			o_rVel:=i_rVel_Film;
		END_IF
	END_IF

	IF NOT i_xAdjustMode THEN(*放牵调整开关@打开了不能使用pid*)
		i_xPidType:=FALSE;
	END_IF

	(*2024.05.25.110051*)
	rTmp:=i_rVel_Film+rYout;
	IF i_xPidType THEN(*放牵使用新方式*)
		o_rVel:=rTmp-rDelt;
		IF o_rVel<0 THEN
			o_rVel:=0;
		END_IF
	ELSE(*原来方式*)
		rDelt:=rTmp-o_rVel;
	END_IF

	IF i_xPidType THEN(*放牵使用新方式*)
		o_rPi_Value:= rYout;
	ELSE
		o_rPi_Value:= rFormulaResult;
	END_IF

	o_rVel:=o_rVel+rPseudoRandomAmplitude_Delta;
	(*2024.12.3.084749 叠加一个速度扰动*)
	o_rVel:=o_rVel+rVel_Disturbance;
	o_rForwardStep:= rForwardStep;

	o_xEno:= TRUE;
	xFilmDecFlag:= FALSE;
ELSE
	o_xEno:= FALSE;
	(*2019.10.12.164013|niu.j|牵引料膜速度减速时加规划，防止速度直接突跳到0*)
	(*2021.2.2.110746 调整了下|Liu.yt*)
	IF NOT xFilmDecFlag  THEN
		lrVel_Acceleration:= UINT_TO_LREAL(i_uiMaxVel_UseCalcAcc)/2/1000.0; (*加速度单位: m/min/ms*)
		xFilmDecFlag:= TRUE;
	END_IF
	IF lrVel_Acceleration<>0 THEN
		lrTempVel:= o_rVel-lrVel_Acceleration * i_iCycleTime_Plc;
	ELSE
		lrTempVel:= i_rVel_Film;
	END_IF

	IF lrTempVel>0 THEN
		o_rVel:= LREAL_TO_REAL(lrTempVel);
	ELSE
		o_rVel:= 0;
		xFilmDecFlag:= FALSE;
	END_IF

	rDelt:=0;
END_IF
rPreFilmVelocity:= i_rVel_Film;

IF i_rUsingGirth<>0 THEN
	o_rVel_rpm:=o_rVel/i_rUsingGirth*1000;(*R/MIN*)
ELSE
	IF i_rGirth_Input<>0 THEN
		o_rVel_rpm:=o_rVel/i_rGirth_Input*1000;(*R/MIN*)
	ELSE
		o_rVel_rpm:=0;(*R/MIN*)
	END_IF
END_IF
o_rVel_rpm:=ABS(o_rVel_rpm);

(* ---- KS_FB_VelocityToVoltage_IfOf.st ---- *)
(*@CES
Name=KS_FB_VelocityToVoltage_IfOf
Type=FunctionBlock
TypeGuid=6f9dac99-8de1-4efc-8465-68ac443b7d08
Guid=4be52c15-88f8-41f0-baca-d2b67222a9df
HasDeclaration=True
HasImplementation=True
*)
{DECLARATION}
FUNCTION_BLOCK KS_FB_VelocityToVoltage_IfOf
VAR_INPUT
	i_xEn: BOOL;
	i_rVel: REAL;
	i_rVel_Film: REAL;
	i_xMachineRev: BOOL;
	i_rUsingGirth: REAL;
	i_rGirth: REAL;
	i_xInchEn: BOOL;
	i_xInchBtn: BOOL;
	i_xInchDir: BOOL;
	i_iInchVel: INT;
	i_iRatedRpm: INT;
	i_iRatedFrq: INT;
	i_iUpperFrq: INT;
	i_uiNum: UINT;
	i_uiDen: UINT;

END_VAR
VAR_OUTPUT
	o_xEn: BOOL;
	o_rVolt: REAL;
	o_rVolt_Film: REAL;
END_VAR
VAR
	rUsingGirth: REAL;
	rRpm_Max: REAL;
	rVel_Max: REAL;
	rVel_Max_Film: REAL;
	rVel_Temp: REAL;
	rFilmVel_Temp: REAL;
END_VAR

{IMPLEMENTATION}
IF i_xEn THEN
	IF i_iRatedRpm<>0 AND i_iRatedFrq<>0 AND
		i_iUpperFrq<>0 AND i_uiNum<>0 AND i_uiDen<>0 THEN
		rUsingGirth:= i_rUsingGirth;
		rRpm_Max:=INT_TO_REAL(i_iUpperFrq)/i_iRatedFrq*i_iRatedRpm;
		rVel_Max:=rRpm_Max*rUsingGirth*i_uiDen/i_uiNum/1000;
		rVel_Max_Film:=rRpm_Max*i_rGirth*i_uiDen/i_uiNum/1000;
		IF i_xMachineRev THEN
			rVel_Temp:= -i_rVel;
			rFilmVel_Temp:= -i_rVel_Film;
		ELSE
			rVel_Temp:= i_rVel;
			rFilmVel_Temp:= i_rVel_Film;
		END_IF
		IF i_xInchEn THEN
			IF i_xInchBtn THEN
				IF i_xInchDir THEN
					rVel_Temp:= -i_iInchVel;
				ELSE
					rVel_Temp:= i_iInchVel;
				END_IF
			END_IF
		END_IF
		IF rVel_Max<>0 THEN
			o_rVolt:= rVel_Temp*10.0/rVel_Max;
		END_IF
		//牵引变频自调
		IF rVel_Max_Film<>0 THEN
			o_rVolt_Film:= rFilmVel_Temp*10.0/rVel_Max_Film;
		END_IF
	ELSE
		o_rVolt:= 0;
		o_rVolt_Film:= 0;
	END_IF
END_IF
